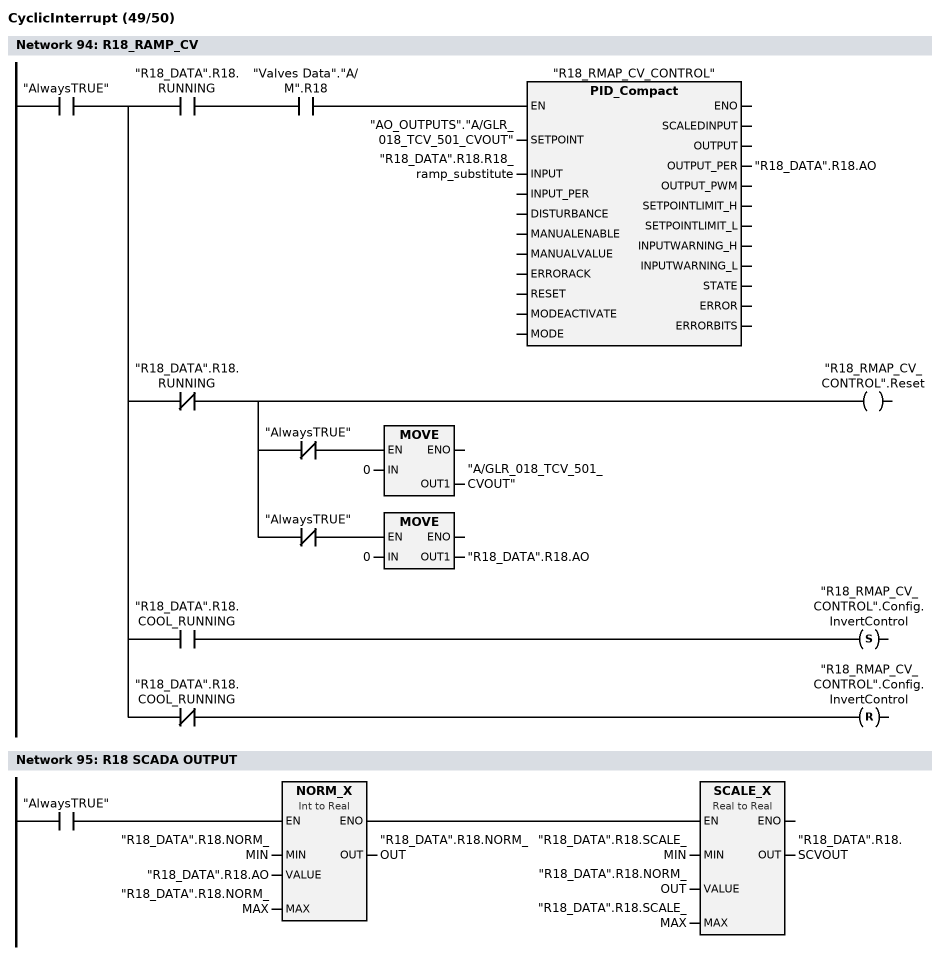
   RUNG wire#powerrail
      Contact( "AlwaysTRUE" )
      wire#w1
      Contact( "R18_DATA".R18.RUNNING )
      Contact( "Valves Data"."A/M".R18 )
      "R18_RMAP_CV_CONTROL".PID_Compact(Setpoint := "AO_OUTPUTS"."A/GLR_018_TCV_501_CVOUT", Input := "R18_DATA".R18.R18_ramp_substitute, Input_PER :=, Disturbance :=, ManualEnable :=, ManualValue :=, ErrorAck :=, Reset :=, ModeActivate :=, Mode :=, ScaledInput =>, Output =>, Output_PER => "R18_DATA".R18.AO, Output_PWM =>, SetpointLimit_H =>, SetpointLimit_L =>, InputWarning_H =>, InputWarning_L =>, State =>, Error =>, ErrorBits =>)
   END_RUNG
   RUNG wire#w1
      I_Contact( "R18_DATA".R18.RUNNING )
      wire#w2
      Coil( "R18_RMAP_CV_CONTROL".Reset )
   END_RUNG
   RUNG wire#w2
      I_Contact( "AlwaysTRUE" )
      Move(in := 0, out1 => "A/GLR_018_TCV_501_CVOUT")
   END_RUNG
   RUNG wire#w2
      I_Contact( "AlwaysTRUE" )
      Move(in := 0, out1 => "R18_DATA".R18.AO)
   END_RUNG
   RUNG wire#w1
      Contact( "R18_DATA".R18.COOL_RUNNING )
      S_Coil( "R18_RMAP_CV_CONTROL".Config.InvertControl )
   END_RUNG
   RUNG wire#w1
      I_Contact( "R18_DATA".R18.COOL_RUNNING )
      R_Coil( "R18_RMAP_CV_CONTROL".Config.InvertControl )
   END_RUNG
   // the same network as SCL:
   #_w1 := "AlwaysTRUE";
   IF "AlwaysTRUE" AND "R18_DATA".R18.RUNNING AND "Valves Data"."A/M".R18 THEN
       "R18_RMAP_CV_CONTROL"(Setpoint := "AO_OUTPUTS"."A/GLR_018_TCV_501_CVOUT",   // PID_Compact
                             Input := "R18_DATA".R18.R18_ramp_substitute,
                             Output_PER => "R18_DATA".R18.AO);
   END_IF;
   "R18_RMAP_CV_CONTROL".Reset := #_w1 AND NOT "R18_DATA".R18.RUNNING;
   IF "R18_RMAP_CV_CONTROL".Reset AND NOT "AlwaysTRUE" THEN
       "A/GLR_018_TCV_501_CVOUT" := 0;
       "R18_DATA".R18.AO := 0;
   END_IF;
   IF #_w1 AND "R18_DATA".R18.COOL_RUNNING THEN "R18_RMAP_CV_CONTROL".Config.InvertControl := TRUE; END_IF;
   IF #_w1 AND NOT "R18_DATA".R18.COOL_RUNNING THEN
       "R18_RMAP_CV_CONTROL".Config.InvertControl := FALSE;
   END_IF;
END_REGION

REGION Network 95: R18 SCADA OUTPUT
   RUNG wire#powerrail
      Contact( "AlwaysTRUE" )
      { S7_Templates := "[SrcType := Int, DestType := Real]" } Normalize(min := "R18_DATA".R18.NORM_MIN, value := "R18_DATA".R18.AO, max := "R18_DATA".R18.NORM_MAX, out => "R18_DATA".R18.NORM_OUT)
      { S7_Templates := "[SrcType := Real, DestType := Real]" } Scale(min := "R18_DATA".R18.SCALE_MIN, value := "R18_DATA".R18.NORM_OUT, max := "R18_DATA".R18.SCALE_MAX, out => "R18_DATA".R18.SCVOUT)
   END_RUNG
   // the same network as SCL:
   IF "AlwaysTRUE" THEN
       "R18_DATA".R18.NORM_OUT := NORM_X(MIN := "R18_DATA".R18.NORM_MIN, VALUE := "R18_DATA".R18.AO, MAX := "R18_DATA".R18.NORM_MAX);
       "R18_DATA".R18.SCVOUT := SCALE_X(MIN := "R18_DATA".R18.SCALE_MIN, VALUE := "R18_DATA".R18.NORM_OUT, MAX := "R18_DATA".R18.SCALE_MAX);
   END_IF;
END_REGION

REGION Network 96: R14 AUTO/MANUAL OUTPUT
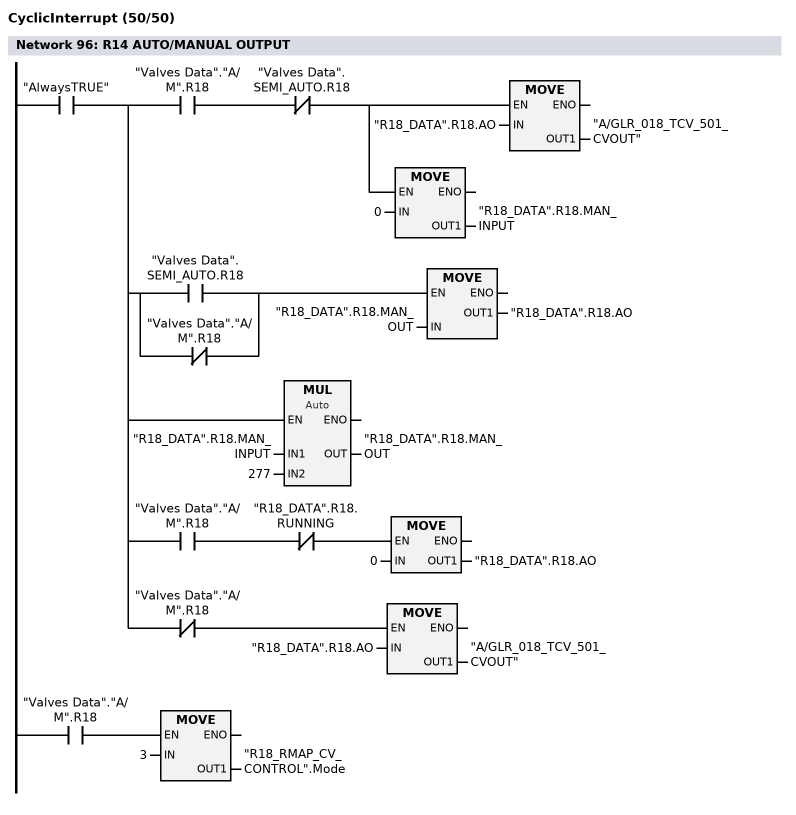
   RUNG wire#powerrail
      Contact( "AlwaysTRUE" )
      wire#w1
      Contact( "Valves Data"."A/M".R18 )
      I_Contact( "Valves Data".SEMI_AUTO.R18 )
      wire#w2
      Move(in := "R18_DATA".R18.AO, out1 => "A/GLR_018_TCV_501_CVOUT")
   END_RUNG
   RUNG wire#w2
      Move(in := 0, out1 => "R18_DATA".R18.MAN_INPUT)
   END_RUNG
   RUNG wire#w1
      Contact( "Valves Data".SEMI_AUTO.R18 )
      wire#w3
      Move(in := "R18_DATA".R18.MAN_OUT, out1 => "R18_DATA".R18.AO)
   END_RUNG
   RUNG wire#w1
      I_Contact( "Valves Data"."A/M".R18 )
   END_RUNG wire#w3
   RUNG wire#w1
      Mul(in1 := "R18_DATA".R18.MAN_INPUT, in2 := 277, out => "R18_DATA".R18.MAN_OUT)
   END_RUNG
   RUNG wire#w1
      Contact( "Valves Data"."A/M".R18 )
      I_Contact( "R18_DATA".R18.RUNNING )
      Move(in := 0, out1 => "R18_DATA".R18.AO)
   END_RUNG
   RUNG wire#w1
      I_Contact( "Valves Data"."A/M".R18 )
      Move(in := "R18_DATA".R18.AO, out1 => "A/GLR_018_TCV_501_CVOUT")
   END_RUNG
   RUNG wire#powerrail
      Contact( "Valves Data"."A/M".R18 )
      Move(in := 3, out1 => "R18_RMAP_CV_CONTROL".Mode)
   END_RUNG
   // the same network as SCL:
   IF "AlwaysTRUE" AND "Valves Data"."A/M".R18 AND NOT "Valves Data".SEMI_AUTO.R18 THEN
       "A/GLR_018_TCV_501_CVOUT" := "R18_DATA".R18.AO;
       "R18_DATA".R18.MAN_INPUT := 0;
   END_IF;
   IF "AlwaysTRUE" AND ("Valves Data".SEMI_AUTO.R18 OR NOT "Valves Data"."A/M".R18) THEN
       "R18_DATA".R18.AO := "R18_DATA".R18.MAN_OUT;
   END_IF;
   IF "AlwaysTRUE" THEN "R18_DATA".R18.MAN_OUT := "R18_DATA".R18.MAN_INPUT * 277; END_IF;
   IF "AlwaysTRUE" AND "Valves Data"."A/M".R18 AND NOT "R18_DATA".R18.RUNNING THEN
       "R18_DATA".R18.AO := 0;
   END_IF;
   IF "AlwaysTRUE" AND NOT "Valves Data"."A/M".R18 THEN
       "A/GLR_018_TCV_501_CVOUT" := "R18_DATA".R18.AO;
   END_IF;
   IF "Valves Data"."A/M".R18 THEN "R18_RMAP_CV_CONTROL".Mode := 3; END_IF;
END_REGION
END_ORGANIZATION_BLOCK
